Staubli VAL3: comment.pgx

public program comment(bool& x_bRefresh)
  local string l_sString
  local bool l_bResult
  local num l_i
  local num l_nIndex
begin
  for l_i = 0 to size(bComment)-1
    if bComment[l_i]
      bComment[l_i]=false
      l_bResult=userPagePrompt("注释：",l_sString)
      if l_bResult
        l_nIndex=nPageIndex*16+l_i
        //Modify by Liu Zhengang 20251103
        switch nSelType
          case 0,1
            if 15<l_nIndex and l_nIndex<96
              call IOcomment(nSelType,l_nIndex,l_sString)
            else
              userPageAlert("此信号不可修改注释！")
            endIf
            io:libSave()
            delay(0.1)
            x_bRefresh=true
          break
          case 2,3
            if 4<l_nIndex and l_nIndex<20
              call IOcomment(nSelType,l_nIndex,l_sString)
            else
              userPageAlert("此信号不可修改注释！")
            endIf
            io:libSave()
            delay(0.1)
            x_bRefresh=true
          break
        endSwitch
      endIf
    endIf
  endFor
end
